// TIA Portal V19 export
// export: Created 2026-10-15T09:44:24.767195Z, ExportSetting WithDefaults, DisplayName Totally Integrated Automation Portal, DisplayVersion V19, DisplayName TIA Portal Openness, DisplayVersion V19, DisplayName TIA Portal Version Control Interface, DisplayVersion V19, DisplayName STEP 7 Professional, DisplayVersion V19, DisplayName STEP 7 Safety, DisplayVersion V19, DisplayName WinCC Basic/Comfort/Advanced, DisplayVersion V19, DisplayName WinCC Unified, DisplayVersion V19
FUNCTION "ROLL_PB21" : Void   // FC29, SCL
{ S7_Optimized_Access := 'TRUE' }
VERSION : 0.1
// stored: AutoNumber true, IsIECCheckEnabled false, SetENOAutomatically false, UDAEnableTagReadback false
   VAR_TEMP
      r : Bool;
      a1 : Word;
      a2 : Word;
      activeDataBlock : Int;
      comparisonResults : Array[0..0] of Bool;
   END_VAR
BEGIN

   #r := FALSE;
   #a1 := W#16#0000;
   #a2 := W#16#0000;
   #activeDataBlock := 0;
   // PB21, STEP 5 network 1
   #activeDataBlock := 15;
   // PB21, STEP 5 network 2
   #r := ((NOT "ROLL_IO".Input[3, 6]) AND (NOT "ROLL_State".M[13, 1]) AND (NOT "ROLL_State".M[5, 6]));
   "ROLL_State".M[99, 7] := #r;
   // PB21, STEP 5 network 3
   #r := ((NOT "ROLL_State".M[13, 3]) AND (NOT "ROLL_State".M[16, 6]) AND (NOT "ROLL_State".M[6, 0]) AND (NOT "ROLL_State".M[6, 2]) AND "ROLL_IO".Input[3, 0] AND "ROLL_IO".Input[5, 0] AND "ROLL_IO".Input[5, 2] AND "ROLL_IO".Input[5, 4]);
   "ROLL_State".M[100, 0] := #r;
   // PB21, STEP 5 network 4
   #r := "ROLL_State".M[190, 6];
   IF #r THEN
       "ROLL_State".M[100, 1] := TRUE;
   END_IF;
   #r := (((NOT "ROLL_State".M[190, 6]) AND "ROLL_IO".Input[5, 3]) OR (NOT "ROLL_IO".Input[0, 1]) OR (NOT "ROLL_State".M[0, 3]) OR (NOT "ROLL_State".M[100, 0]) OR "ROLL_State".M[190, 5]);
   IF #r THEN
       "ROLL_State".M[100, 1] := FALSE;
   END_IF;
   // PB21, STEP 5 network 5
   #r := "ROLL_State".M[190, 6];
   IF #r THEN
       "ROLL_State".M[100, 2] := TRUE;
   END_IF;
   #r := (("ROLL_IO".Input[5, 3] AND "ROLL_IO".Input[5, 6]) OR (NOT "ROLL_IO".Input[0, 1]) OR (NOT "ROLL_State".M[0, 3]) OR (NOT "ROLL_State".M[100, 0]) OR "ROLL_State".M[190, 5]);
   IF #r THEN
       "ROLL_State".M[100, 2] := FALSE;
   END_IF;
   // PB21, STEP 5 network 6
   #r := "ROLL_State".M[190, 6];
   IF #r THEN
       "ROLL_State".M[100, 3] := TRUE;
   END_IF;
   #r := (((NOT "ROLL_IO".Input[7, 5]) AND (NOT "ROLL_State".M[190, 6])) OR (NOT "ROLL_IO".Input[0, 1]) OR (NOT "ROLL_State".M[0, 3]) OR (NOT "ROLL_State".M[100, 0]) OR "ROLL_State".M[190, 5] OR "ROLL_State".M[5, 6] OR "ROLL_State".M[8, 5]);
   IF #r THEN
       "ROLL_State".M[100, 3] := FALSE;
   END_IF;
   // PB21, STEP 5 network 7
   #r := "ROLL_State".M[190, 6];
   IF #r THEN
       "ROLL_State".M[100, 4] := TRUE;
   END_IF;
   #r := (((NOT "ROLL_State".M[100, 0]) AND (NOT "ROLL_State".M[190, 6])) OR (NOT "ROLL_IO".Input[0, 1]) OR (NOT "ROLL_State".M[0, 3]) OR (NOT "ROLL_State".M[99, 7]) OR "ROLL_State".M[190, 5]);
   IF #r THEN
       "ROLL_State".M[100, 4] := FALSE;
   END_IF;
   // PB21, STEP 5 network 8
   #r := ((NOT "ROLL_State".M[31, 5]) AND (NOT "ROLL_State".M[5, 6]) AND ((NOT "ROLL_IO".Input[5, 6]) OR (NOT "ROLL_State".S5Timers[70].Q)) AND "ROLL_IO".Input[0, 2] AND "ROLL_IO".Input[3, 1] AND "ROLL_State".M[100, 0]);
   "ROLL_State".M[100, 5] := #r;
   // PB21, STEP 5 network 9
   #r := ((("ROLL_IO".Input[7, 5] AND "ROLL_State".S5Timers[97].Q) OR (NOT "ROLL_State".S5Timers[96].Q)) AND "ROLL_State".M[0, 3] AND "ROLL_State".M[100, 5]);
   "ROLL_State".M[100, 6] := #r;
   // PB21, STEP 5 network 10
   #r := ((((NOT "ROLL_IO".Input[7, 5]) AND "ROLL_State".S5Timers[96].Q) OR (NOT "ROLL_State".S5Timers[97].Q)) AND "ROLL_State".M[0, 3] AND "ROLL_State".M[100, 5]);
   "ROLL_State".M[100, 7] := #r;
   // PB21, STEP 5 network 11
   #r := "ROLL_State".M[190, 6];
   IF #r THEN
       "ROLL_State".M[101, 1] := TRUE;
   END_IF;
   #r := (((NOT "ROLL_State".M[190, 6]) AND "ROLL_IO".Input[5, 3] AND "ROLL_IO".Input[5, 6] AND "ROLL_IO".Input[6, 0]) OR (NOT "ROLL_IO".Input[0, 1]) OR (NOT "ROLL_State".M[0, 3]) OR (NOT "ROLL_State".M[100, 0]) OR "ROLL_State".M[190, 5]);
   IF #r THEN
       "ROLL_State".M[101, 1] := FALSE;
   END_IF;
   // PB21, STEP 5 network 12
   #r := "ROLL_State".M[190, 6];
   IF #r THEN
       "ROLL_State".M[101, 2] := TRUE;
   END_IF;
   #r := (((NOT "ROLL_State".M[190, 6]) AND "ROLL_IO".Input[5, 3] AND "ROLL_IO".Input[5, 6] AND "ROLL_IO".Input[6, 0]) OR (NOT "ROLL_IO".Input[0, 1]) OR (NOT "ROLL_State".M[0, 3]) OR (NOT "ROLL_State".M[100, 0]) OR "ROLL_State".M[190, 5]);
   IF #r THEN
       "ROLL_State".M[101, 2] := FALSE;
   END_IF;
   // PB21, STEP 5 network 13
   #r := "ROLL_State".M[190, 6];
   IF #r THEN
       "ROLL_State".M[101, 3] := TRUE;
   END_IF;
   #r := (((NOT "ROLL_State".M[190, 6]) AND ((NOT "ROLL_IO".Input[7, 5]) OR "ROLL_IO".Input[6, 0])) OR (NOT "ROLL_IO".Input[0, 1]) OR (NOT "ROLL_State".M[0, 3]) OR (NOT "ROLL_State".M[100, 0]) OR "ROLL_State".M[190, 5] OR "ROLL_State".M[5, 6] OR "ROLL_State".M[8, 5]);
   IF #r THEN
       "ROLL_State".M[101, 3] := FALSE;
   END_IF;
   // PB21, STEP 5 network 14
   #r := "ROLL_State".M[190, 6];
   IF #r THEN
       "ROLL_State".M[101, 4] := TRUE;
   END_IF;
   #r := (((NOT "ROLL_State".M[190, 6]) AND "ROLL_IO".Input[6, 0]) OR (NOT "ROLL_IO".Input[0, 1]) OR (NOT "ROLL_State".M[0, 3]) OR (NOT "ROLL_State".M[100, 0]) OR (NOT "ROLL_State".M[99, 7]) OR "ROLL_State".M[190, 5]);
   IF #r THEN
       "ROLL_State".M[101, 4] := FALSE;
   END_IF;
   // PB21, STEP 5 network 15
   #a2 := #a1;
   #a1 := W#16#2005;
   #r := "ROLL_IO".Input[6, 0];
   "ROLL_TimerOp"(Number := 121,
                  Operation := 0,
                  Signal := #r,
                  Preset := #a1);
   // PB21, STEP 5 network 16
   #r := ((NOT "ROLL_State".M[31, 5]) AND (NOT "ROLL_State".M[5, 6]) AND (((NOT "ROLL_State".S5Timers[121].Q) AND "ROLL_State".M[101, 5]) OR (NOT "ROLL_IO".Input[6, 0])) AND "ROLL_IO".Input[0, 2] AND "ROLL_IO".Input[3, 1] AND "ROLL_State".M[100, 0]);
   "ROLL_State".M[101, 5] := #r;
   // PB21, STEP 5 network 17
   #r := ((("ROLL_IO".Input[7, 5] AND "ROLL_State".S5Timers[97].Q) OR (NOT "ROLL_State".S5Timers[96].Q)) AND "ROLL_State".M[101, 5]);
   "ROLL_State".M[101, 6] := #r;
   // PB21, STEP 5 network 18
   #r := ((((NOT "ROLL_IO".Input[7, 5]) AND "ROLL_State".S5Timers[96].Q) OR (NOT "ROLL_State".S5Timers[97].Q)) AND "ROLL_State".M[101, 5]);
   "ROLL_State".M[101, 7] := #r;
   // PB21, STEP 5 network 19
   #r := "ROLL_State".M[190, 6];
   IF #r THEN
       "ROLL_State".M[102, 1] := TRUE;
   END_IF;
   #r := (((NOT "ROLL_State".M[190, 6]) AND "ROLL_IO".Input[5, 3] AND "ROLL_IO".Input[5, 6] AND "ROLL_IO".Input[6, 0] AND "ROLL_IO".Input[6, 2]) OR (NOT "ROLL_IO".Input[0, 1]) OR (NOT "ROLL_State".M[0, 3]) OR (NOT "ROLL_State".M[100, 0]) OR "ROLL_State".M[190, 5]);
   IF #r THEN
       "ROLL_State".M[102, 1] := FALSE;
   END_IF;
   // PB21, STEP 5 network 20
   #r := "ROLL_State".M[190, 6];
   IF #r THEN
       "ROLL_State".M[102, 2] := TRUE;
   END_IF;
   #r := (((NOT "ROLL_State".M[190, 6]) AND "ROLL_IO".Input[6, 2]) OR (NOT "ROLL_IO".Input[0, 1]) OR (NOT "ROLL_State".M[0, 3]) OR (NOT "ROLL_State".M[100, 0]) OR "ROLL_State".M[190, 5]);
   IF #r THEN
       "ROLL_State".M[102, 2] := FALSE;
   END_IF;
   // PB21, STEP 5 network 21
   #r := "ROLL_State".M[190, 6];
   IF #r THEN
       "ROLL_State".M[102, 3] := TRUE;
   END_IF;
   #r := (((NOT "ROLL_State".M[190, 6]) AND ((NOT "ROLL_IO".Input[7, 5]) OR "ROLL_IO".Input[6, 2])) OR (NOT "ROLL_IO".Input[0, 1]) OR (NOT "ROLL_State".M[0, 3]) OR (NOT "ROLL_State".M[100, 0]) OR "ROLL_State".M[190, 5] OR "ROLL_State".M[5, 6] OR "ROLL_State".M[8, 5]);
   IF #r THEN
       "ROLL_State".M[102, 3] := FALSE;
   END_IF;
   // PB21, STEP 5 network 22
   #r := "ROLL_State".M[190, 6];
   IF #r THEN
       "ROLL_State".M[102, 4] := TRUE;
   END_IF;
   #r := (((NOT "ROLL_State".M[190, 6]) AND "ROLL_IO".Input[6, 2]) OR (NOT "ROLL_IO".Input[0, 1]) OR (NOT "ROLL_State".M[0, 3]) OR (NOT "ROLL_State".M[100, 0]) OR (NOT "ROLL_State".M[99, 7]) OR "ROLL_State".M[190, 5]);
   IF #r THEN
       "ROLL_State".M[102, 4] := FALSE;
   END_IF;
   // PB21, STEP 5 network 23
   #r := ((NOT "ROLL_State".M[31, 5]) AND (NOT "ROLL_State".M[5, 6]) AND (NOT "ROLL_State".S5Timers[72].Q) AND "ROLL_IO".Input[0, 2] AND "ROLL_IO".Input[3, 1] AND "ROLL_State".M[100, 0]);
   "ROLL_State".M[102, 5] := #r;
   // PB21, STEP 5 network 24
   #r := ((("ROLL_IO".Input[7, 5] AND "ROLL_State".S5Timers[97].Q) OR (NOT "ROLL_State".S5Timers[96].Q)) AND "ROLL_State".M[0, 3] AND "ROLL_State".M[102, 5]);
   "ROLL_State".M[102, 6] := #r;
   // PB21, STEP 5 network 25
   #r := ((((NOT "ROLL_IO".Input[7, 5]) AND "ROLL_State".S5Timers[96].Q) OR (NOT "ROLL_State".S5Timers[97].Q) OR "ROLL_State".M[0, 4]) AND "ROLL_State".M[102, 5]);
   "ROLL_State".M[102, 7] := #r;
   // PB21, STEP 5 network 26
   #r := "ROLL_State".M[190, 6];
   IF #r THEN
       "ROLL_State".M[105, 1] := TRUE;
   END_IF;
   #r := (((NOT "ROLL_State".M[190, 6]) AND "ROLL_State".M[0, 4]) OR (NOT "ROLL_IO".Input[0, 1]) OR (NOT "ROLL_State".M[0, 3]) OR (NOT "ROLL_State".M[100, 0]) OR "ROLL_State".M[190, 5]);
   IF #r THEN
       "ROLL_State".M[105, 1] := FALSE;
   END_IF;
   // PB21, STEP 5 network 27
   #r := "ROLL_State".M[190, 6];
   IF #r THEN
       "ROLL_State".M[105, 2] := TRUE;
   END_IF;
   #r := ((NOT "ROLL_IO".Input[0, 1]) OR (NOT "ROLL_State".M[0, 3]) OR (NOT "ROLL_State".M[100, 0]) OR "ROLL_IO".Input[6, 2] OR "ROLL_State".M[190, 5]);
   IF #r THEN
       "ROLL_State".M[105, 2] := FALSE;
   END_IF;
   // PB21, STEP 5 network 28
   #r := "ROLL_State".M[190, 6];
   IF #r THEN
       "ROLL_State".M[105, 3] := TRUE;
   END_IF;
   #r := (((NOT "ROLL_State".M[190, 6]) AND ((NOT "ROLL_IO".Input[7, 5]) OR "ROLL_State".M[0, 4])) OR (NOT "ROLL_IO".Input[0, 1]) OR (NOT "ROLL_State".M[0, 3]) OR (NOT "ROLL_State".M[100, 0]) OR "ROLL_State".M[190, 5] OR "ROLL_State".M[5, 6] OR "ROLL_State".M[8, 5]);
   IF #r THEN
       "ROLL_State".M[105, 3] := FALSE;
   END_IF;
   // PB21, STEP 5 network 29
   #r := "ROLL_State".M[190, 6];
   IF #r THEN
       "ROLL_State".M[105, 4] := TRUE;
   END_IF;
   #r := (((NOT "ROLL_State".M[190, 6]) AND "ROLL_State".M[0, 4]) OR (NOT "ROLL_IO".Input[0, 1]) OR (NOT "ROLL_State".M[0, 3]) OR (NOT "ROLL_State".M[100, 0]) OR (NOT "ROLL_State".M[99, 7]) OR "ROLL_State".M[190, 5]);
   IF #r THEN
       "ROLL_State".M[105, 4] := FALSE;
   END_IF;
   // PB21, STEP 5 network 30
   #a2 := #a1;
   #a1 := W#16#2005;
   #r := "ROLL_State".M[0, 4];
   "ROLL_TimerOp"(Number := 120,
                  Operation := 0,
                  Signal := #r,
                  Preset := #a1);
   // PB21, STEP 5 network 31
   #r := ((NOT "ROLL_State".M[31, 5]) AND (NOT "ROLL_State".M[5, 6]) AND (((NOT "ROLL_State".S5Timers[120].Q) AND "ROLL_State".M[105, 5]) OR (NOT "ROLL_State".M[0, 4])) AND "ROLL_IO".Input[0, 2] AND "ROLL_IO".Input[3, 1] AND "ROLL_State".M[100, 0]);
   "ROLL_State".M[105, 5] := #r;
   // PB21, STEP 5 network 32
   #r := ((("ROLL_IO".Input[7, 5] AND "ROLL_State".S5Timers[97].Q) OR (NOT "ROLL_State".S5Timers[96].Q)) AND "ROLL_State".M[105, 5]);
   "ROLL_State".M[105, 6] := #r;
   // PB21, STEP 5 network 33
   #r := ((((NOT "ROLL_IO".Input[7, 5]) AND "ROLL_State".S5Timers[96].Q) OR (NOT "ROLL_State".S5Timers[97].Q)) AND "ROLL_State".M[105, 5]);
   "ROLL_State".M[105, 7] := #r;
   // PB21, STEP 5 network 34
   #r := ((((NOT "ROLL_IO".Input[5, 5]) AND ("ROLL_State".M[40, 5] OR "ROLL_State".M[42, 1]) AND "ROLL_State".M[31, 5]) OR (NOT "ROLL_IO".Input[5, 6])) AND "ROLL_IO".Input[0, 2] AND "ROLL_IO".Input[3, 1] AND "ROLL_State".M[100, 0]);
   "ROLL_State".M[103, 0] := #r;
   // PB21, STEP 5 network 35
   #r := (((NOT "ROLL_IO".Input[5, 3]) OR (NOT "ROLL_IO".Input[6, 0]) OR (NOT "ROLL_State".S5Timers[121].Q)) AND "ROLL_IO".Input[3, 1] AND "ROLL_State".M[100, 0] AND "ROLL_State".M[31, 5]);
   "ROLL_State".M[103, 3] := #r;
   // PB21, STEP 5 network 36
   #r := (((NOT "ROLL_IO".Input[5, 6]) AND "ROLL_IO".Input[0, 2]) OR (("ROLL_State".M[103, 0] OR "ROLL_State".M[103, 3]) AND "ROLL_State".S5Timers[62].Q AND "ROLL_State".S5Timers[97].Q));
   "ROLL_State".M[103, 1] := #r;
   // PB21, STEP 5 network 37
   #r := ((NOT "ROLL_IO".Input[6, 2]) AND "ROLL_IO".Input[3, 1] AND "ROLL_State".M[100, 0] AND "ROLL_State".M[31, 5]);
   "ROLL_State".M[103, 4] := #r;
   // PB21, STEP 5 network 38
   #a2 := #a1;
   #a1 := W#16#1050;
   #r := ("ROLL_IO".Output[22, 3] AND "ROLL_State".M[103, 4]);
   "ROLL_TimerOp"(Number := 119,
                  Operation := 1,
                  Signal := #r,
                  Preset := #a1);
   // PB21, STEP 5 network 39
   #r := (((("ROLL_State".M[103, 0] OR "ROLL_State".M[103, 3]) AND "ROLL_State".S5Timers[96].Q) OR "ROLL_State".M[103, 4] OR "ROLL_State".S5Timers[119].Q) AND "ROLL_State".S5Timers[62].Q);
   "ROLL_State".M[103, 2] := #r;
   // PB21, STEP 5 network 40
   #r := "ROLL_State".M[190, 6];
   IF #r THEN
       "ROLL_State".M[104, 0] := TRUE;
   END_IF;
   #r := (((NOT "ROLL_State".M[190, 6]) AND ((NOT "ROLL_IO".Input[5, 0]) OR (NOT "ROLL_IO".Input[5, 2]) OR (NOT "ROLL_IO".Input[5, 4]))) OR (NOT "ROLL_IO".Input[0, 1]) OR (NOT "ROLL_IO".Input[7, 0]) OR (NOT "ROLL_State".M[26, 5]) OR (NOT "ROLL_State".M[99, 7]) OR "ROLL_State".M[16, 6] OR "ROLL_State".M[190, 5]);
   IF #r THEN
       "ROLL_State".M[104, 0] := FALSE;
   END_IF;
   // PB21, STEP 5 network 41
   #r := "ROLL_State".M[190, 6];
   IF #r THEN
       "ROLL_State".M[104, 1] := TRUE;
   END_IF;
   #r := (((NOT "ROLL_State".M[190, 6]) AND ((NOT "ROLL_IO".Input[5, 0]) OR (NOT "ROLL_IO".Input[5, 2]) OR (NOT "ROLL_IO".Input[5, 4]))) OR (NOT "ROLL_IO".Input[0, 1]) OR (NOT "ROLL_State".M[26, 0]) OR (NOT "ROLL_State".M[99, 7]) OR "ROLL_State".M[16, 6] OR "ROLL_State".M[190, 5]);
   IF #r THEN
       "ROLL_State".M[104, 1] := FALSE;
   END_IF;
   // PB21, STEP 5 network 42
   #r := "ROLL_State".M[190, 6];
   IF #r THEN
       "ROLL_State".M[104, 4] := TRUE;
   END_IF;
   #r := (((NOT "ROLL_State".M[190, 6]) AND ((NOT "ROLL_IO".Input[5, 0]) OR (NOT "ROLL_IO".Input[5, 2]) OR (NOT "ROLL_IO".Input[5, 4]))) OR (NOT "ROLL_IO".Input[0, 1]) OR (NOT "ROLL_IO".Input[4, 7]) OR (NOT "ROLL_State".M[27, 4]) OR (NOT "ROLL_State".M[99, 7]) OR "ROLL_State".M[16, 6] OR "ROLL_State".M[190, 5]);
   IF #r THEN
       "ROLL_State".M[104, 4] := FALSE;
   END_IF;
   // PB21, STEP 5 network 43
   #r := "ROLL_State".M[190, 6];
   IF #r THEN
       "ROLL_State".M[104, 5] := TRUE;
   END_IF;
   #r := (((NOT "ROLL_State".M[190, 6]) AND "ROLL_IO".Input[5, 3] AND "ROLL_IO".Input[5, 6] AND "ROLL_IO".Input[6, 0] AND "ROLL_IO".Input[6, 2]) OR (NOT "ROLL_IO".Input[0, 1]) OR (NOT "ROLL_State".M[100, 0]) OR (NOT "ROLL_State".M[24, 1]) OR "ROLL_State".M[190, 5]);
   IF #r THEN
       "ROLL_State".M[104, 5] := FALSE;
   END_IF;
   // PB21, STEP 5 network 44
   #r := "ROLL_State".M[190, 6];
   IF #r THEN
       "ROLL_State".M[104, 6] := TRUE;
   END_IF;
   #r := (((NOT "ROLL_State".M[190, 6]) AND (("ROLL_IO".Input[5, 3] AND "ROLL_IO".Input[5, 6] AND "ROLL_IO".Input[6, 0]) OR (NOT "ROLL_IO".Input[7, 5]))) OR (NOT "ROLL_IO".Input[0, 1]) OR (NOT "ROLL_State".M[100, 0]) OR (NOT "ROLL_State".M[25, 0]) OR "ROLL_State".M[190, 5] OR "ROLL_State".M[5, 6] OR "ROLL_State".M[8, 5]);
   IF #r THEN
       "ROLL_State".M[104, 6] := FALSE;
   END_IF;
   // PB21, STEP 5 network 45
   #r := "ROLL_State".S5Timers[59].Q;
   "ROLL_IO".Output[17, 0] := #r;
   // PB21, STEP 5 network 46
   #r := ("ROLL_IO".Input[6, 5] AND "ROLL_State".M[100, 0]);
   "ROLL_IO".Output[17, 5] := #r;
   RETURN;
END_FUNCTION
